// TIA Portal V20 export
Screen "190J5RoofGeo"  1276x673
  ScreenItem "permanentareaborderrectangle" at 0,0 size 0x0  Type=HmiRectangle
  ScreenItem "Button_Back" at 2,2 size 90x60  Type=HmiButton
  ScreenItem "Move_Legend" at 1182,2 size 90x60  Type=HmiButton
  ScreenItem "Fusszeile_Button_ManualOPMode1_2" at 279,2 size 90x60  Type=HmiButton
  ScreenItem "面板容器_2" at 1090,4 size 88x58  Type=HmiFaceplateContainer
  ScreenItem "OPMode1_Blocked" at 1164,6 size 14x14  Type=HmiGraphicView
  ScreenItem "OPMode4_Foreground_Blocked" at 1089,5 size 88x58  Type=HmiGraphicView
  ScreenItem "Fusszeile_Button_ManualOPMode1_1" at 95,2 size 90x60  Type=HmiButton
  ScreenItem "Button_Back_1" at 1180,606 size 90x60  Type=HmiButton
  ScreenItem "Fusszeile_Button_ManualOPMode1_3" at 187,2 size 90x60  Type=HmiButton
  ScreenItem "Fusszeile_Button_ManualOPMode1_4" at 997,2 size 90x60  Type=HmiButton
  ScreenItem "Fusszeile_Button_ManualOPMode1_5" at 902,1 size 90x60  Type=HmiButton
  ScreenItem "文本域_14" at 936,-172 size 140x40  Type=HmiTextBox
  ScreenItem "Title_ScreenOverview_X390_Y2_1" at 384,5 size 510x57  Type=HmiTextBox
  ScreenItem "Graphic view_1" at 195,176 size 864x387  Type=HmiGraphicView
  ScreenItem "Line_Header_X0_Y64" at -3,67 size 1276x0  Type=HmiLine
  ScreenItem "Rectangle_1" at 0,0 size 152x48  Type=HmiRectangle
  ScreenItem "文本域_11" at 2,1 size 122x45  Type=HmiTextBox
  ScreenItem "圆_1" at 0,0 size 100x30  Type=HmiCircle
  ScreenItem "圆_2" at 0,0 size 100x30  Type=HmiCircle
  ScreenItem "Rectangle_2" at 0,0 size 152x48  Type=HmiRectangle
  ScreenItem "文本域_1" at 2,1 size 122x45  Type=HmiTextBox
  ScreenItem "圆_3" at 0,0 size 100x30  Type=HmiCircle
  ScreenItem "圆_4" at 0,0 size 100x30  Type=HmiCircle
  ScreenItem "Rectangle_3" at 0,0 size 152x48  Type=HmiRectangle
  ScreenItem "文本域_2" at 2,1 size 122x45  Type=HmiTextBox
  ScreenItem "圆_5" at 0,0 size 100x30  Type=HmiCircle
  ScreenItem "圆_6" at 0,0 size 100x30  Type=HmiCircle
